Fanuc KAREL source: kf00082.KL

-- PROVISIONAL review KL for V770-1; original PC SHA256 9a230a3c923e7d13ceb0ec02ed8f431b75f6cd90f3cfc03fa2316d8f9fcb875a
-- Incomplete behavior may be omitted. Consult companion uncertainty JSON. Do not deploy.
PROGRAM KF00082
%NOLOCKGROUP
BEGIN
  -- UNRESOLVED_PC offsets 5-15; opcodes 27,22,31
  -- UNRESOLVED_PC offsets 20-54; opcodes 27,27,2E,22,22,22,22,31
  -- UNRESOLVED_PC offsets 59-93; opcodes 27,22,22,22,22,22,31
  -- UNRESOLVED_PC offsets 98-102; opcodes 7F
END KF00082
